FUNCTION_BLOCK NOOP_INIT (* No-Op, auch bekannt als "No Operation" mit INIT - wrapt NOOP, reicht INIT direkt auf INITO durch *)
  (* Standard: 61131-3; Classification: standard boolean function; Description: Copyright (c) 2026 Meisterschulen am Ostbahnhof This program and the accompanying materials are made available under the terms of the Eclipse Public License 2.0 which is available at https://www.eclipse.org/legal/epl-2.0/ SPDX-License-Identifier: EPL-2.0 *)
  (* Version 1.1, 2026-10-11, Franz Höpfinger, Meisterschulen am Ostbahnhof, Copyright-Header, Classification und Remarks nachgezogen; Doku ergaenzt. Interne Umsetzung wrapt jetzt NOOP statt iec61131::selection::F_MOVE - damit entfaellt dieser iec61131-3-Abhaengigkeitspfad. *)
  (* Version 1.0, 2026-05-05, franz, Meisterschulen am Ostbahnhof, initial API and implementation and/or initial documentation *)
  PACKAGE iec61131::booleanOperators;
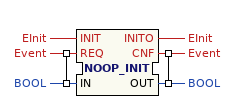
  EVENT_INPUT
    INIT : EInit; (* Initialization Request *)
    REQ WITH IN; (* Normal Execution Request *)
  END_EVENT
  EVENT_OUTPUT
    INITO : EInit; (* Initialization Confirm *)
    CNF WITH OUT; (* Execution Confirmation *)
  END_EVENT
  VAR_INPUT
    IN : BOOL; (* Input *)
  END_VAR
  VAR_OUTPUT
    OUT : BOOL; (* Output *)
  END_VAR
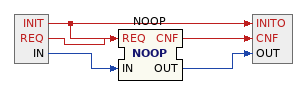
  FBS
    NOOP : iec61131::booleanOperators::NOOP;
  END_FBS
  EVENT_CONNECTIONS
    INIT TO INITO;
    INIT TO NOOP.REQ;
    REQ TO NOOP.REQ;
    NOOP.CNF TO CNF;
  END_CONNECTIONS
  DATA_CONNECTIONS
    IN TO NOOP.IN;
    NOOP.OUT TO OUT;
  END_CONNECTIONS
END_FUNCTION_BLOCK
